FUNCTION_BLOCK running_version
  VAR
  END_VAR
  VAR_INPUT
    s1 : BOOL;
    s2 : BOOL;
    reset : BOOL;
  END_VAR
  VAR_OUTPUT
    k1 : BOOL;
    k2 : BOOL;
  END_VAR

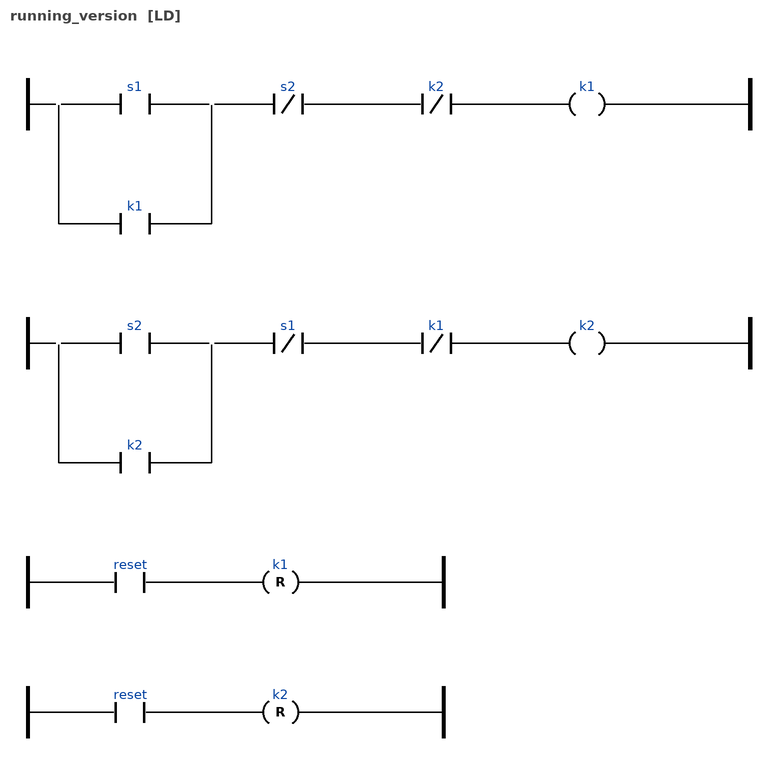
(* LD diagram, written out as Structured Text *)
k1 := (s1 OR k1) AND NOT s2 AND NOT k2;
k2 := (s2 OR k2) AND NOT s1 AND NOT k1;
IF reset THEN k1 := FALSE; END_IF;
IF reset THEN k2 := FALSE; END_IF;
END_FUNCTION_BLOCK
